VAR_GLOBAL
{IF defined (S85_HW)}
    bWorkshopMainButton AT %I* : BOOL;
    bWorkshopMainLightRelay AT %Q* : BOOL;
{END_IF}
END_VAR

(* stored: Version 1.1.0.1
   GVL GVL_BeckhoffIO: Id {9dbe3bca-c820-4c58-b452-4f0928e0acb4} *)
